Fanuc KAREL source: kb00197.compact.KL

PROGRAM KB00197
%STACKSIZE=65535
%PRIORITY=65535
%NOLOCKGROUP
VAR
P1 : FILE
P2 : STRING[80]
P3 : INTEGER
P4 : INTEGER
BEGIN
P2='A'
P3=1
P4=1
WRITE_DICT(P1,P2,P3,P4)
END KB00197
